PROGRAM MAIN
VAR_INPUT
END_VAR
VAR_OUTPUT
END_VAR
VAR
	fHysteresis: REAL := 1;
	fbSR: SR;
END_VAR
VAR // added by the converter: edge detectors and wires of the graphical bodies
    _w1 : REAL;
    _w2, _w4 : ANY;
    _w3 : BOOL;
END_VAR

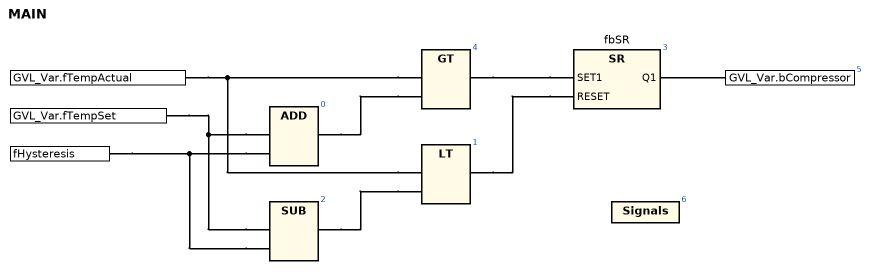
_w1 := GVL_Var.fTempSet + fHysteresis;
_w3 := GVL_Var.fTempActual < _w2;
_w2 := GVL_Var.fTempSet - fHysteresis;
fbSR(SET1 := _w4, RESET := _w3); // SR
_w4 := GVL_Var.fTempActual > _w1;
GVL_Var.bCompressor := fbSR.Q1;
Signals();

END_PROGRAM

(* stored: Version 1.1.0.1, ProductVersion 3.1.4024.16
   POU MAIN: Id {b541f825-9a7d-4070-85a6-a54fc02dbf05}, SpecialFunc None *)
